// SIMATIC S7-200 SMART project (STEP 7-Micro/WIN SMART), CPU SR30

SYMBOL_TABLE STATES
ONSTATE          M0.0     // SYSTEM ON
CONVEYOR_RUN_STATE M0.1     // CONVEYOR ON
CONVEYOR_CW_STATE M0.2     // COUNTERCLOCKWISE STATE
ACTUATOR_ON_STATE M0.3     // ACTUATOR STATE ON
PROCESS_STATE    M0.4     // PROCESSING
ENTER_STATE      M0.5     // ENTER PROTECTION
RED_GOT_REJECTED M0.6     // RED_GOT_REJECTED
WHITE_GOT_REJECTED M0.7     // WHITE_GOT_REJECTED
END_SYMBOL_TABLE

SYMBOL_TABLE SET
WHITE_SELECTED   M2.1     // WHITE SET PRIORITY
RED_SELECTED     M2.0     // RED SET PRIORITY
COLOR_SELECTED   M2.2     // COLOR HAS BEEN SELECTED
END_SYMBOL_TABLE

SYMBOL_TABLE TIMERS
TIMER_WHITE      T32      // TIMER
TIMER_RED        T33      // TIMER RED
END_SYMBOL_TABLE

SYMBOL_TABLE System Symbols_0
Always_On        SM0.0    // Always ON
END_SYMBOL_TABLE

SYMBOL_TABLE HMI_INPUTS
WHITE_PRIORITY   M1.1     // WHITE ONLY
RED_PRIORITY     M1.0     // RED ONLY
HMI_STOP         M1.3     // HMI STOP
HMI_START        M1.2     // HMI START
HMI_RESET        M1.4     // HMI RESET
HMI_PAUSE        M1.6     // HMI PAUSE
HMI_ENTER_BUTTON M1.5     // HMI ENTER BUTTON FOR PRIORITY LIMIT
END_SYMBOL_TABLE

SYMBOL_TABLE COMMUNICATION
COMMMUNICATION   V100.5   // COMMUNICATION
MASTER_START     V101.5   // MASTER_START
MASTER_STOP      V102.5   // MASTER_STOP
MASTER_RESET     V103.5   // MASTER_RESET
END_SYMBOL_TABLE

SYMBOL_TABLE ANALOG VALUES
CONVERTED_LIMIT  VW3000   // LIMIT IN PLC ALREADY
HMI_INSERT_LIMIT VW500    // HMI_Counter_Limit
REJECTED_COUNTER C0       // REJECTED_COUNTER
END_SYMBOL_TABLE

SYMBOL_TABLE HMI INDICATORS
ONLINE_LED       M3.0     // ONLINE_LED
PROCESS_LED      M3.1     // PROCESS_LED
HALTED_LED       M3.2     // HALTED_LED
READY_LED        M3.3     // READY_LED
COMMUNICATION_LED M3.4     // COMMUNICATION_LED
MOTOR_LED        M3.5     // MOTOR LED
ALARM            M3.6     // ALARM SET OFF
END_SYMBOL_TABLE

ORGANIZATION_BLOCK MAIN:OB1
TITLE=Program Comments
BEGIN
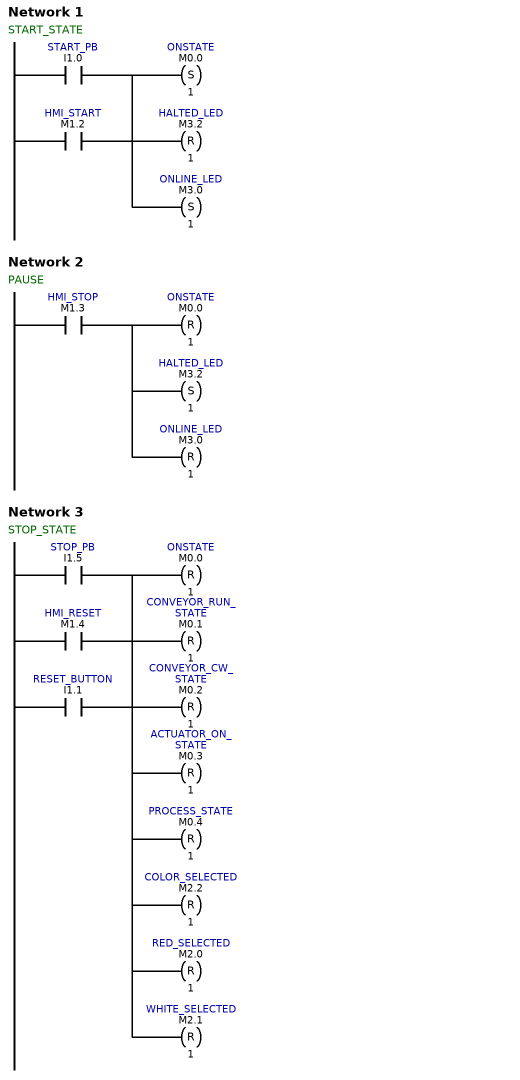
Network 1
// START_STATE
LD     START_PB:I1.0
O      HMI_START:M1.2
S      ONSTATE:M0.0, 1
R      HALTED_LED:M3.2, 1
S      ONLINE_LED:M3.0, 1
Network 2
// PAUSE
LD     HMI_STOP:M1.3
R      ONSTATE:M0.0, 1
S      HALTED_LED:M3.2, 1
R      ONLINE_LED:M3.0, 1
Network 3
// STOP_STATE
LD     STOP_PB:I1.5
O      HMI_RESET:M1.4
O      RESET_BUTTON:I1.1
R      ONSTATE:M0.0, 1
R      CONVEYOR_RUN_STATE:M0.1, 1
R      CONVEYOR_CW_STATE:M0.2, 1
R      ACTUATOR_ON_STATE:M0.3, 1
R      PROCESS_STATE:M0.4, 1
R      COLOR_SELECTED:M2.2, 1
R      RED_SELECTED:M2.0, 1
R      WHITE_SELECTED:M2.1, 1
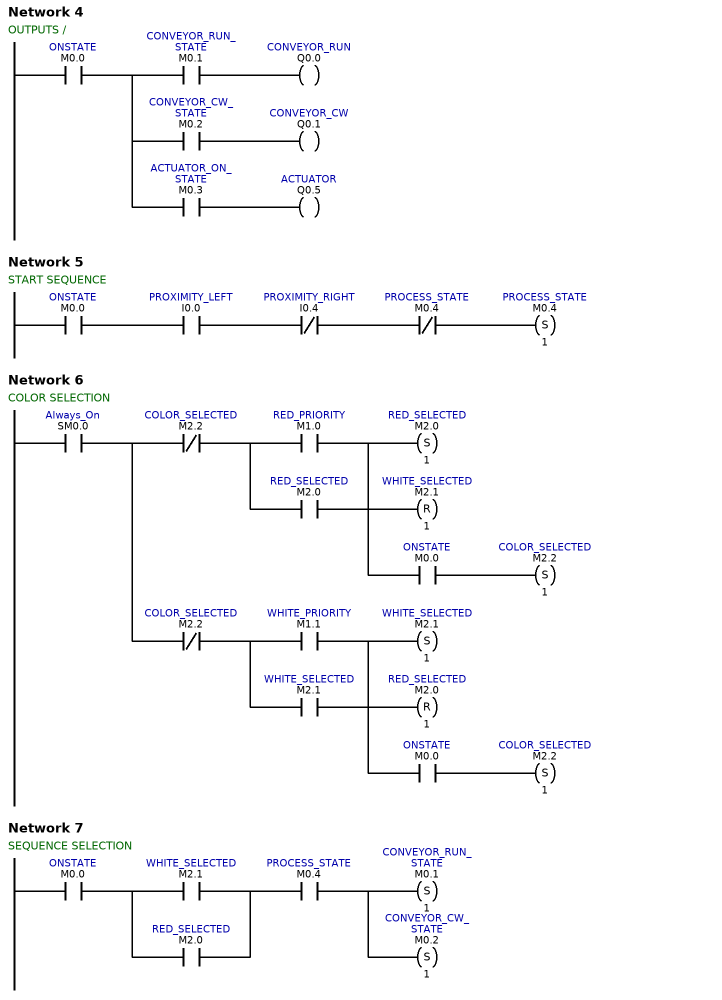
Network 4
// OUTPUTS
// 
LD     ONSTATE:M0.0
LPS
A      CONVEYOR_RUN_STATE:M0.1
=      CONVEYOR_RUN:Q0.0
LRD
A      CONVEYOR_CW_STATE:M0.2
=      CONVEYOR_CW:Q0.1
LPP
A      ACTUATOR_ON_STATE:M0.3
=      ACTUATOR:Q0.5
Network 5
// START SEQUENCE
LD     ONSTATE:M0.0
A      PROXIMITY_LEFT:I0.0
AN     PROXIMITY_RIGHT:I0.4
AN     PROCESS_STATE:M0.4
S      PROCESS_STATE:M0.4, 1
Network 6
// COLOR SELECTION
LD     Always_On:SM0.0
LPS
AN     COLOR_SELECTED:M2.2
LD     RED_PRIORITY:M1.0
O      RED_SELECTED:M2.0
ALD
S      RED_SELECTED:M2.0, 1
R      WHITE_SELECTED:M2.1, 1
A      ONSTATE:M0.0
S      COLOR_SELECTED:M2.2, 1
LPP
AN     COLOR_SELECTED:M2.2
LD     WHITE_PRIORITY:M1.1
O      WHITE_SELECTED:M2.1
ALD
S      WHITE_SELECTED:M2.1, 1
R      RED_SELECTED:M2.0, 1
A      ONSTATE:M0.0
S      COLOR_SELECTED:M2.2, 1
Network 7
// SEQUENCE SELECTION
LD     ONSTATE:M0.0
LD     WHITE_SELECTED:M2.1
O      RED_SELECTED:M2.0
ALD
A      PROCESS_STATE:M0.4
S      CONVEYOR_RUN_STATE:M0.1, 1
S      CONVEYOR_CW_STATE:M0.2, 1
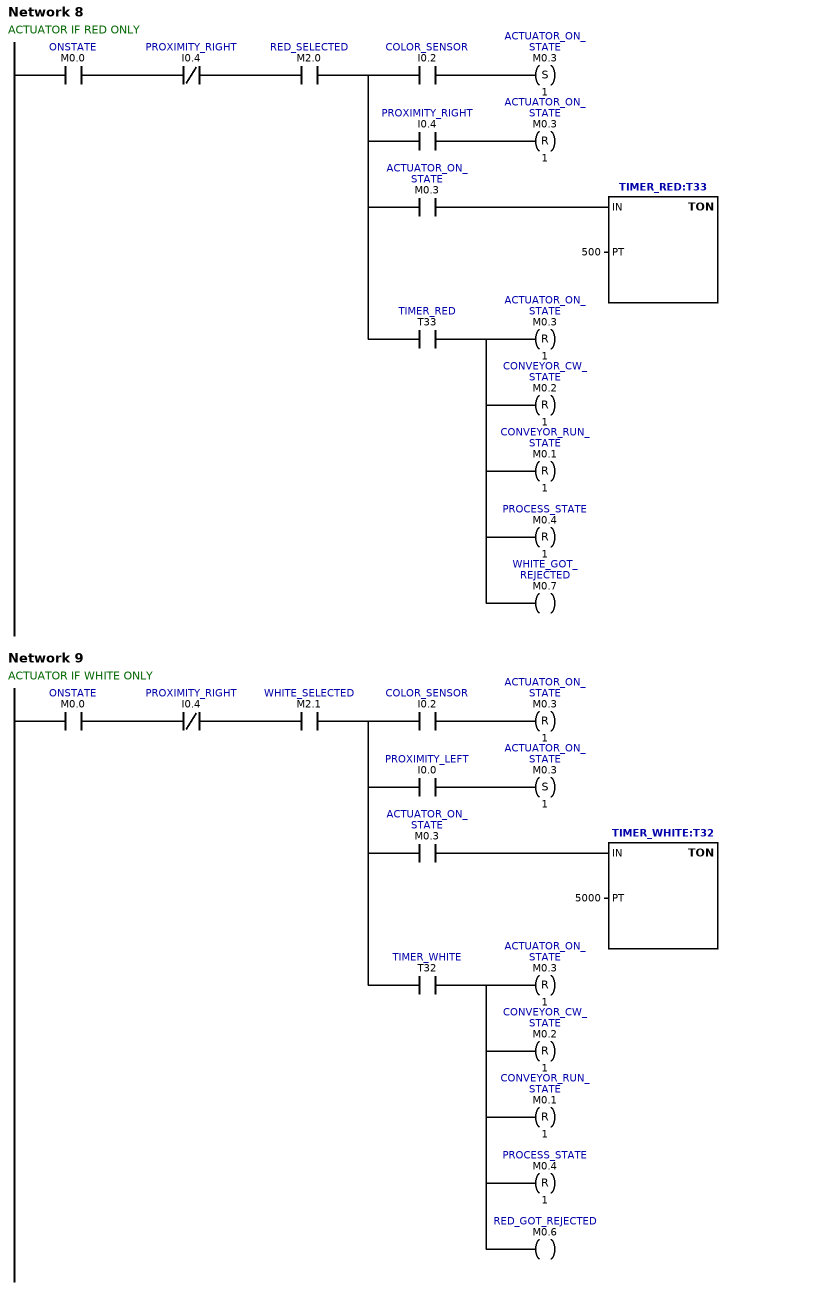
Network 8
// ACTUATOR IF RED ONLY
LD     ONSTATE:M0.0
AN     PROXIMITY_RIGHT:I0.4
A      RED_SELECTED:M2.0
LPS
A      COLOR_SENSOR:I0.2
S      ACTUATOR_ON_STATE:M0.3, 1
LRD
A      PROXIMITY_RIGHT:I0.4
R      ACTUATOR_ON_STATE:M0.3, 1
LRD
A      ACTUATOR_ON_STATE:M0.3
TON    TIMER_RED:T33, 500
LPP
A      TIMER_RED:T33
R      ACTUATOR_ON_STATE:M0.3, 1
R      CONVEYOR_CW_STATE:M0.2, 1
R      CONVEYOR_RUN_STATE:M0.1, 1
R      PROCESS_STATE:M0.4, 1
=      WHITE_GOT_REJECTED:M0.7
Network 9
// ACTUATOR IF WHITE ONLY
LD     ONSTATE:M0.0
AN     PROXIMITY_RIGHT:I0.4
A      WHITE_SELECTED:M2.1
LPS
A      COLOR_SENSOR:I0.2
R      ACTUATOR_ON_STATE:M0.3, 1
LRD
A      PROXIMITY_LEFT:I0.0
S      ACTUATOR_ON_STATE:M0.3, 1
LRD
A      ACTUATOR_ON_STATE:M0.3
TON    TIMER_WHITE:T32, 5000
LPP
A      TIMER_WHITE:T32
R      ACTUATOR_ON_STATE:M0.3, 1
R      CONVEYOR_CW_STATE:M0.2, 1
R      CONVEYOR_RUN_STATE:M0.1, 1
R      PROCESS_STATE:M0.4, 1
=      RED_GOT_REJECTED:M0.6
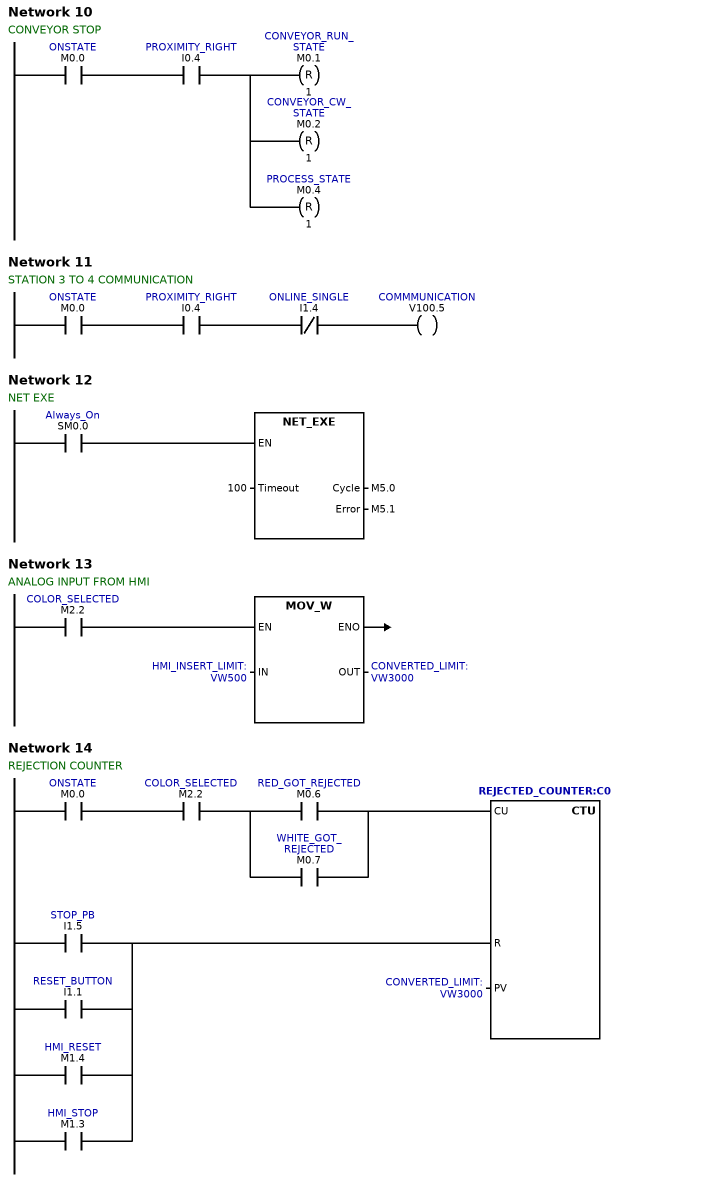
Network 10
// CONVEYOR STOP
LD     ONSTATE:M0.0
A      PROXIMITY_RIGHT:I0.4
R      CONVEYOR_RUN_STATE:M0.1, 1
R      CONVEYOR_CW_STATE:M0.2, 1
R      PROCESS_STATE:M0.4, 1
Network 11
// STATION 3 TO 4 COMMUNICATION
LD     ONSTATE:M0.0
A      PROXIMITY_RIGHT:I0.4
AN     ONLINE_SINGLE:I1.4
=      COMMMUNICATION:V100.5
Network 12
// NET EXE
LD     Always_On:SM0.0
CALL   NET_EXE:SBR1, 100, M5.0, M5.1
Network 13
// ANALOG INPUT FROM HMI
LD     COLOR_SELECTED:M2.2
MOVW   HMI_INSERT_LIMIT:VW500, CONVERTED_LIMIT:VW3000
Network 14
// REJECTION COUNTER
LD     ONSTATE:M0.0
A      COLOR_SELECTED:M2.2
LD     RED_GOT_REJECTED:M0.6
O      WHITE_GOT_REJECTED:M0.7
ALD
LD     STOP_PB:I1.5
O      RESET_BUTTON:I1.1
O      HMI_RESET:M1.4
O      HMI_STOP:M1.3
CTU    REJECTED_COUNTER:C0, CONVERTED_LIMIT:VW3000
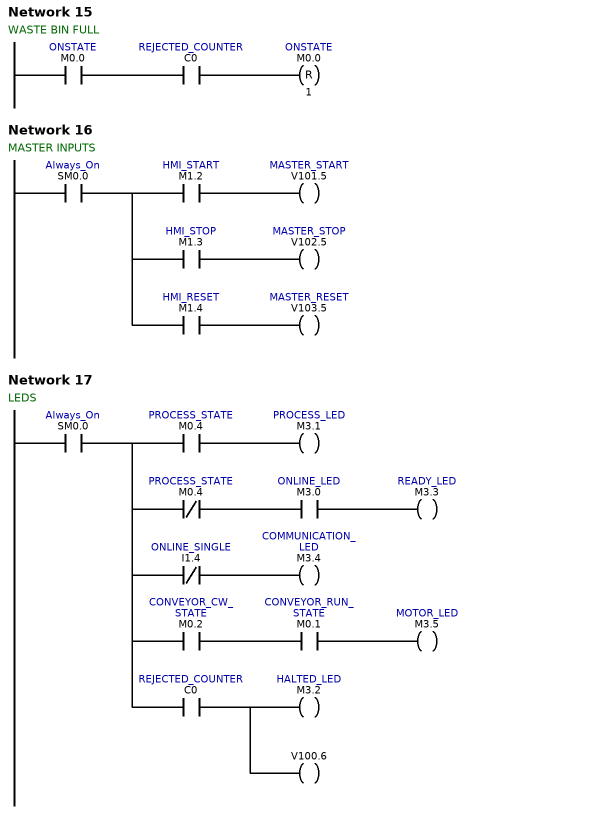
Network 15
// WASTE BIN FULL
LD     ONSTATE:M0.0
A      REJECTED_COUNTER:C0
R      ONSTATE:M0.0, 1
Network 16
// MASTER INPUTS
LD     Always_On:SM0.0
LPS
A      HMI_START:M1.2
=      MASTER_START:V101.5
LRD
A      HMI_STOP:M1.3
=      MASTER_STOP:V102.5
LPP
A      HMI_RESET:M1.4
=      MASTER_RESET:V103.5
Network 17
// LEDS
LD     Always_On:SM0.0
LPS
A      PROCESS_STATE:M0.4
=      PROCESS_LED:M3.1
LRD
AN     PROCESS_STATE:M0.4
A      ONLINE_LED:M3.0
=      READY_LED:M3.3
LRD
AN     ONLINE_SINGLE:I1.4
=      COMMUNICATION_LED:M3.4
LRD
A      CONVEYOR_CW_STATE:M0.2
A      CONVEYOR_RUN_STATE:M0.1
=      MOTOR_LED:M3.5
LPP
A      REJECTED_COUNTER:C0
=      HALTED_LED:M3.2
=      V100.6
END_ORGANIZATION_BLOCK

// SBR1: protected block, not included
